(* IEC 61131-3 sources: nautilus/examples/it-rack/live, 1 file *)

(* ---- hw_types.st ---- *)
(*
  Generated by `naut snmp import`: the IT-hardware UDT set from
  docs/design/it-drivers.md §2. Do not edit — every importer (snmp, redfish,
  prometheus) writes this same file, so re-running any of them restores it.
  Member order is the wire order the drivers deliver; the compiled TYPE
  must match it slot for slot, which is why it is generated and not typed.
*)

TYPE
  Fan : STRUCT
    Name : STRING;
    Present : BOOL;
    RPM : REAL;
    Pct : REAL;
    Fault : BOOL;
  END_STRUCT;
  PDU : STRUCT
    Online : BOOL;
    Name : STRING;
    Model : STRING;
    Serial : STRING;
    Amps : REAL;
    Watts : REAL;
    Overload : BOOL;
    OutletCount : DINT;
  END_STRUCT;
  PDUOutlet : STRUCT
    Index : DINT;
    Name : STRING;
    On : BOOL;
    Amps : REAL;
    Watts : REAL;
  END_STRUCT;
  PSU : STRUCT
    Name : STRING;
    Present : BOOL;
    Fault : BOOL;
    InputOk : BOOL;
    InputV : REAL;
    OutputW : REAL;
    CapacityW : REAL;
  END_STRUCT;
  Server : STRUCT
    Online : BOOL;
    PowerOn : BOOL;
    Health : DINT;
    Fault : BOOL;
    Warning : BOOL;
    Model : STRING;
    Serial : STRING;
    UptimeS : DINT;
    CpuPct : REAL;
    MemPct : REAL;
    Load1 : REAL;
    RootDiskPct : REAL;
    InletTempC : REAL;
    MaxTempC : REAL;
    PowerW : REAL;
    FanCount : DINT;
    PsuCount : DINT;
    TempCount : DINT;
  END_STRUCT;
  Switch : STRUCT
    Online : BOOL;
    Name : STRING;
    Model : STRING;
    Serial : STRING;
    UptimeS : DINT;
    CpuPct : REAL;
    MemPct : REAL;
    TempC : REAL;
    Fault : BOOL;
    PortsTotal : DINT;
    PortsUp : DINT;
  END_STRUCT;
  SwitchPort : STRUCT
    Index : DINT;
    Name : STRING;
    Alias : STRING;
    AdminUp : BOOL;
    OperUp : BOOL;
    Down : BOOL;
    SpeedMbps : REAL;
    InBps : REAL;
    OutBps : REAL;
    InPct : REAL;
    OutPct : REAL;
    InErrors : DINT;
    OutErrors : DINT;
    InDiscards : DINT;
    OutDiscards : DINT;
    ErrorRate : REAL;
    PoeOn : BOOL;
    PoeW : REAL;
  END_STRUCT;
  TempSensor : STRUCT
    Name : STRING;
    Value : REAL;
    Fault : BOOL;
    High : BOOL;
    HighHigh : BOOL;
    HighSP : REAL;
    HighHighSP : REAL;
  END_STRUCT;
  UPS : STRUCT
    Online : BOOL;
    Name : STRING;
    Model : STRING;
    Serial : STRING;
    OnBattery : BOOL;
    LowBattery : BOOL;
    BatteryFault : BOOL;
    Fault : BOOL;
    ChargePct : REAL;
    RuntimeMin : REAL;
    LoadPct : REAL;
    InputV : REAL;
    OutputV : REAL;
    BatteryTempC : REAL;
  END_STRUCT;
END_TYPE
